(* IEC 61131-3 sources: rusty/tests/lit/cfc/variables/expression_source, 1 file *)

(* ---- main.st ---- *)
FUNCTION main : DINT
    expression_source();
    // CHECK: sum = 4, scaled = -2, ready = 1, idle = 0, differs = 1
    printf('sum = %d, scaled = %d, ready = %d, idle = %d, differs = %d$N', expression_source.sum, expression_source.scaled, expression_source.ready, expression_source.idle, expression_source.differs);

    // `item` reads arr[2] before the last sink overwrites it with `a`.
    // CHECK: item = 30, arr[2] = 3
    printf('item = %d, arr[2] = %d$N', expression_source.item, expression_source.arr[2]);

    // `grid[1, 2]` is written through `grid[i, i + 1]`, then read back doubled.
    // CHECK: grid[1, 2] = 3, cell = 6
    printf('grid[1, 2] = %d, cell = %d$N', expression_source.grid[1, 2], expression_source.cell);
END_FUNCTION
